SUBAPPLICATION GreenWhiteBackground_Auseinanderklappen (* Subapplication Type *)
  (* Standard: 61499-2 *)
  (* Version 1.0, 2023-02-11, franz *)
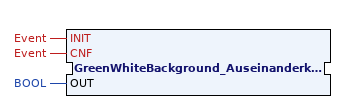
  EVENT_INPUT
    INIT;
    CNF;
  END_EVENT
  VAR_INPUT
    OUT : BOOL;
  END_VAR
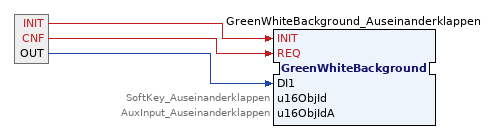
  SUBAPPS
    GreenWhiteBackground_Auseinanderklappen : GreenWhiteBackground(u16ObjId := SoftKey_Auseinanderklappen, u16ObjIdA := AuxInput_Auseinanderklappen);
  END_SUBAPPS
  EVENT_CONNECTIONS
    INIT TO GreenWhiteBackground_Auseinanderklappen.INIT;
    CNF TO GreenWhiteBackground_Auseinanderklappen.REQ;
  END_CONNECTIONS
  DATA_CONNECTIONS
    OUT TO GreenWhiteBackground_Auseinanderklappen.DI1;
  END_CONNECTIONS
END_SUBAPPLICATION
